PROGRAM ControlFBD
VAR
	qxLampStarted	AT %Q* : BOOL;
	qxSliderAout 	AT %Q* : BOOL; 
	qxSliderAin 	AT %Q* : BOOL; 
	qxSliderBout 	AT %Q* : BOOL; 
	qxSliderBin 	AT %Q* : BOOL; 
	qxDrillDown 	AT %Q* : BOOL;
	qxDrillUp		AT %Q* : BOOL;
	qxLampEmStopOk	AT %Q* : BOOL;
	qxLampSafetyOk  AT %Q* : BOOL;
	qxLampHomePos   AT %Q* : BOOL;
	
	
	mxManualRun : BOOL;
	mxEmergencyButtonPressed: BOOL;
	mxAuto : BOOL;
	mxAutoAIn : BOOL;
	mxAutoAOut : BOOL;
	mxAutoBIn : BOOL;
	mxAutoBOut : BOOL;
	mxAutoDrillDown: BOOL;
	mxAutoDrillUp: BOOL;
	
	mxSafetyOK : BOOL;
	mxManualOk : BOOL;
	mxCycleStopActivated : BOOL;
	mxBlink : BOOL;
	
	fbBlink : BLINK;

	
	
	ixButtonStart	AT %I* : BOOL;
	ixButtonStop	AT %I* : BOOL;
	ixSliderAout	AT %I* : BOOL;
	ixSliderAin		AT %I* : BOOL;
	ixSliderBout	AT %I* : BOOL;
	ixSliderBin		AT %I* : BOOL;
	ixDrillUp		AT %I* : BOOL;
	ixDrillDown		AT %I* : BOOL;

	ixAuto			AT %I* : BOOL;
	ixBtn1EmStopOk	AT %I* : BOOL;
	ixBtn2EmStopOk	AT %I* : BOOL;	
	ixSafety1StopOk	AT %I* : BOOL;
	ixSafety2StopOk	AT %I* : BOOL;	
	ixBtnReset		AT %I* : BOOL;
	ixBtnAout		AT %I* : BOOL;
	ixBtnAin		AT %I* : BOOL;
	ixBtnBout		AT %I* : BOOL;
	ixBtnBin		AT %I* : BOOL;
	ixBtnDrillOut	AT %I* : BOOL;
	ixBtnDrillIn	AT %I* : BOOL;

	mx: BOOL;
	mxStart: BOOL;
END_VAR

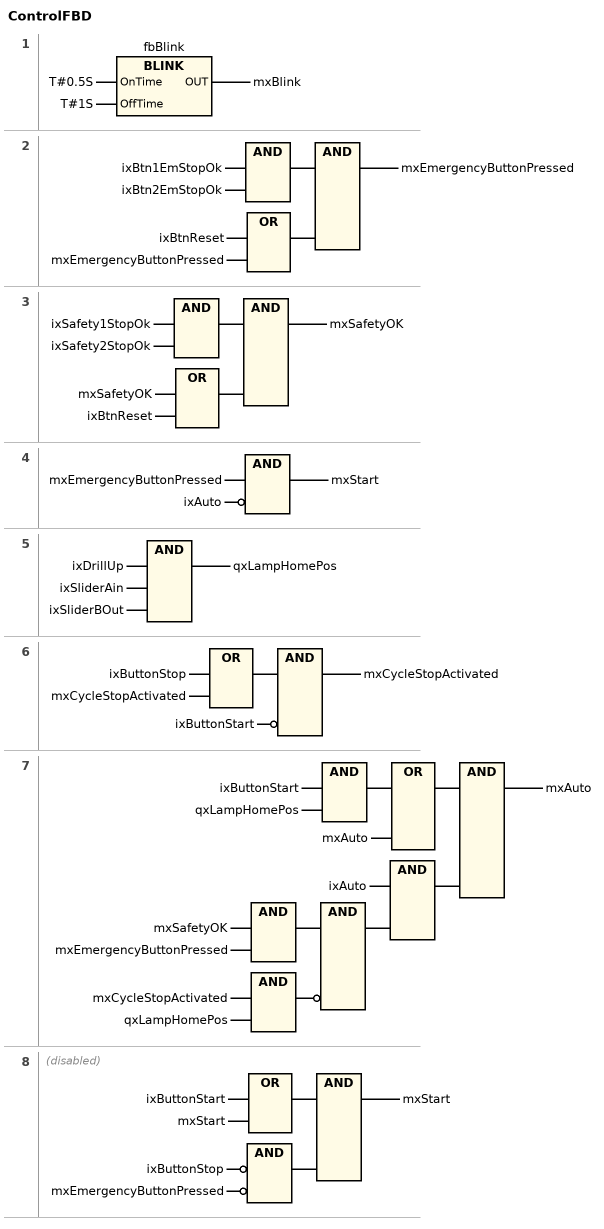
// NETWORK 1
fbBlink(OnTime := T#0.5S, OffTime := T#1S); // BLINK
mxBlink := fbBlink.OUT;

// NETWORK 2
mxEmergencyButtonPressed := (ixBtn1EmStopOk AND ixBtn2EmStopOk) AND (ixBtnReset OR mxEmergencyButtonPressed);

// NETWORK 3
mxSafetyOK := (ixSafety1StopOk AND ixSafety2StopOk) AND (mxSafetyOK OR ixBtnReset);

// NETWORK 4
mxStart := mxEmergencyButtonPressed AND NOT ixAuto;

// NETWORK 5
qxLampHomePos := ixDrillUp AND ixSliderAin AND ixSliderBOut;

// NETWORK 6
mxCycleStopActivated := (ixButtonStop OR mxCycleStopActivated) AND NOT ixButtonStart;

// NETWORK 7
mxAuto := (ixButtonStart AND qxLampHomePos OR mxAuto) AND (ixAuto AND ((mxSafetyOK AND mxEmergencyButtonPressed) AND NOT (mxCycleStopActivated AND qxLampHomePos)));

// NETWORK 8 (disabled)
// mxStart := (ixButtonStart OR mxStart) AND (NOT ixButtonStop AND NOT mxEmergencyButtonPressed);

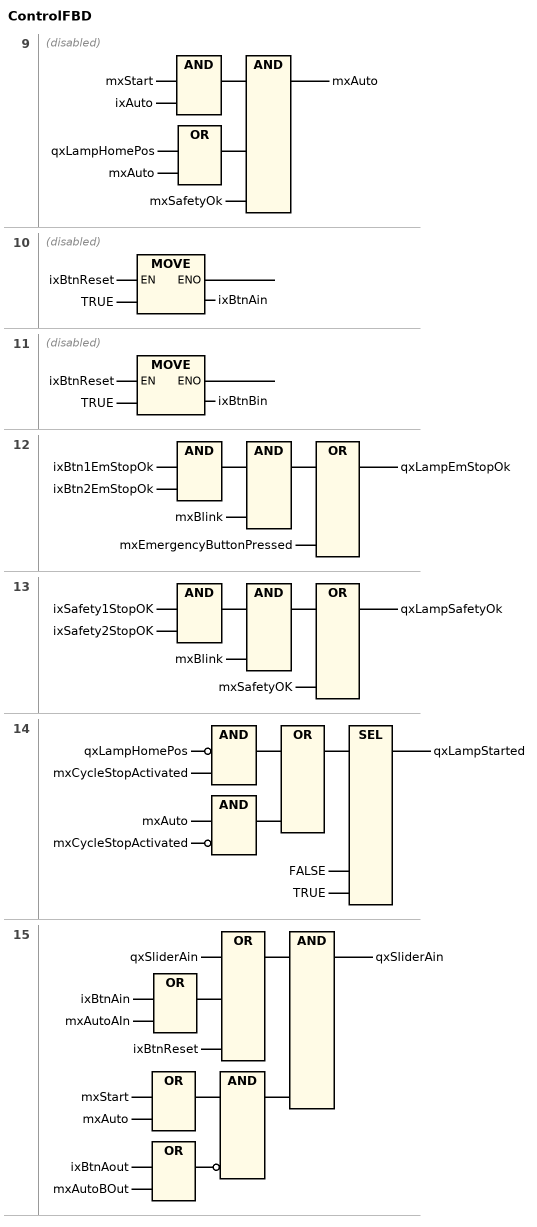
// NETWORK 9 (disabled)
// mxAuto := (mxStart AND ixAuto) AND (qxLampHomePos OR mxAuto) AND mxSafetyOk;

// NETWORK 10 (disabled)
// IF ixBtnReset THEN ixBtnAin := TRUE; END_IF

// NETWORK 11 (disabled)
// IF ixBtnReset THEN ixBtnBin := TRUE; END_IF

// NETWORK 12
qxLampEmStopOk := (ixBtn1EmStopOk AND ixBtn2EmStopOk) AND mxBlink OR mxEmergencyButtonPressed;

// NETWORK 13
qxLampSafetyOk := (ixSafety1StopOK AND ixSafety2StopOK) AND mxBlink OR mxSafetyOK;

// NETWORK 14
qxLampStarted := SEL(NOT qxLampHomePos AND mxCycleStopActivated OR mxAuto AND NOT mxCycleStopActivated, FALSE, TRUE);

// NETWORK 15
qxSliderAin := (qxSliderAin OR (ixBtnAin OR mxAutoAIn) OR ixBtnReset) AND ((mxStart OR mxAuto) AND NOT (ixBtnAout OR mxAutoBOut));

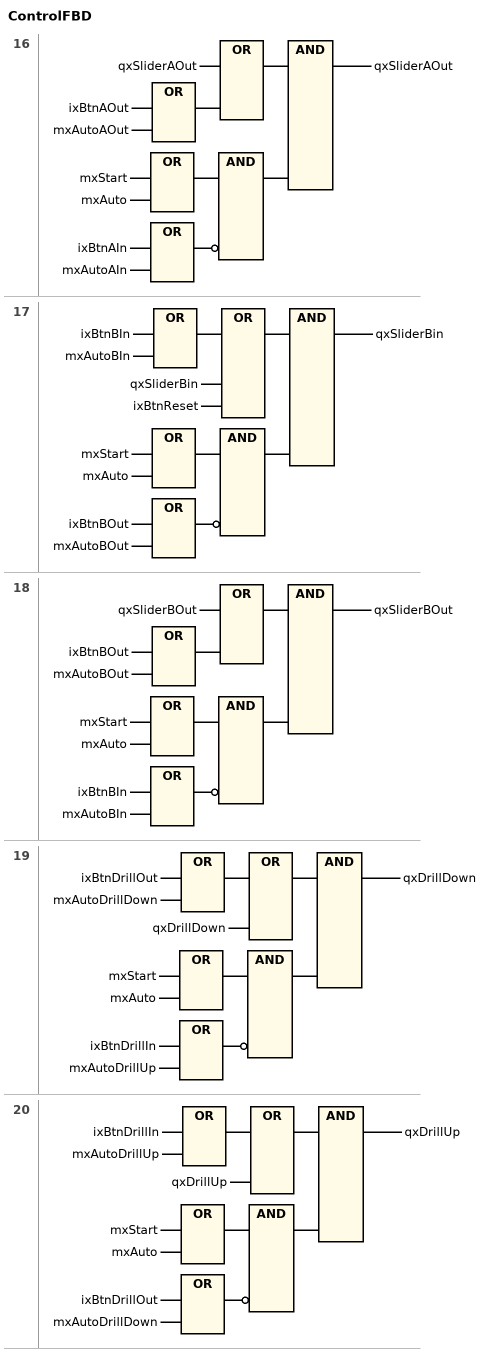
// NETWORK 16
qxSliderAOut := (qxSliderAOut OR (ixBtnAOut OR mxAutoAOut)) AND ((mxStart OR mxAuto) AND NOT (ixBtnAIn OR mxAutoAIn));

// NETWORK 17
qxSliderBin := ((ixBtnBIn OR mxAutoBIn) OR qxSliderBin OR ixBtnReset) AND ((mxStart OR mxAuto) AND NOT (ixBtnBOut OR mxAutoBOut));

// NETWORK 18
qxSliderBOut := (qxSliderBOut OR (ixBtnBOut OR mxAutoBOut)) AND ((mxStart OR mxAuto) AND NOT (ixBtnBIn OR mxAutoBIn));

// NETWORK 19
qxDrillDown := ((ixBtnDrillOut OR mxAutoDrillDown) OR qxDrillDown) AND ((mxStart OR mxAuto) AND NOT (ixBtnDrillIn OR mxAutoDrillUp));

// NETWORK 20
qxDrillUp := ((ixBtnDrillIn OR mxAutoDrillUp) OR qxDrillUp) AND ((mxStart OR mxAuto) AND NOT (ixBtnDrillOut OR mxAutoDrillDown));

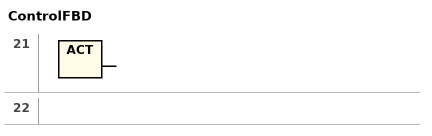
// NETWORK 21
ACT();

// NETWORK 22

ACTION ACT:
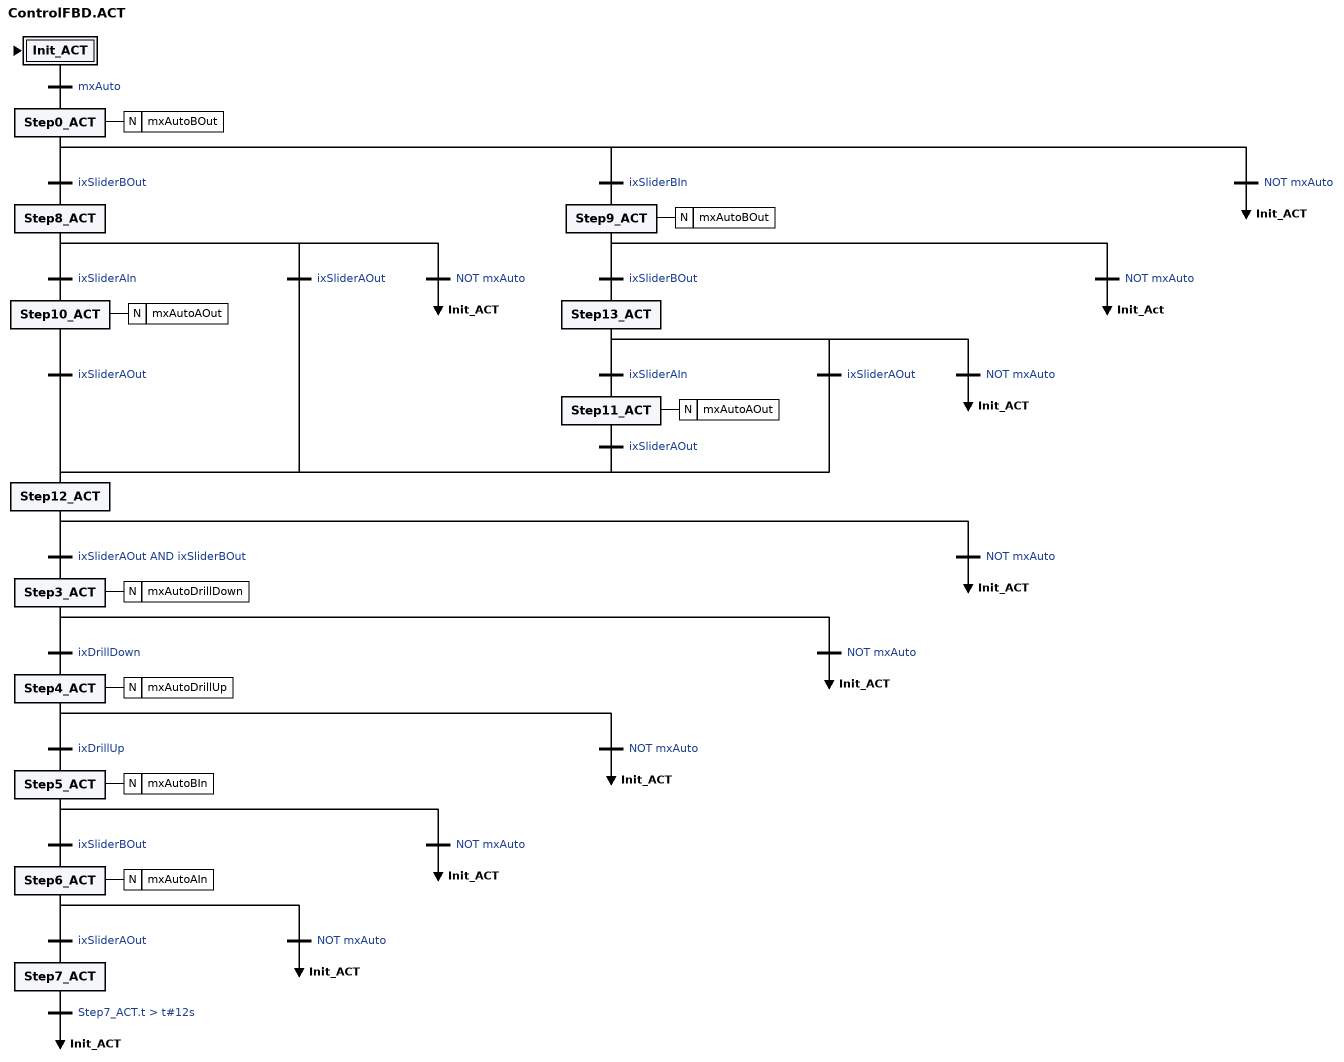
INITIAL_STEP Init_ACT:
END_STEP
TRANSITION FROM Init_ACT TO Step0_ACT
    := mxAuto;
END_TRANSITION
STEP Step0_ACT:
    mxAutoBOut(N);
END_STEP
TRANSITION FROM Step0_ACT TO Step8_ACT
    := ixSliderBOut;
END_TRANSITION
STEP Step8_ACT:
END_STEP
TRANSITION FROM Step8_ACT TO Step10_ACT
    := ixSliderAIn;
END_TRANSITION
STEP Step10_ACT:
    mxAutoAOut(N);
END_STEP
TRANSITION FROM Step10_ACT TO Step12_ACT
    := ixSliderAOut;
END_TRANSITION
TRANSITION FROM Step8_ACT TO Step12_ACT
    := ixSliderAOut;
END_TRANSITION
TRANSITION FROM Step8_ACT TO Init_ACT
    := NOT mxAuto;
END_TRANSITION
TRANSITION FROM Step0_ACT TO Step9_ACT
    := ixSliderBIn;
END_TRANSITION
STEP Step9_ACT:
    mxAutoBOut(N);
END_STEP
TRANSITION FROM Step9_ACT TO Step13_ACT
    := ixSliderBOut;
END_TRANSITION
TRANSITION FROM Step9_ACT TO Init_Act
    := NOT mxAuto;
END_TRANSITION
STEP Step13_ACT:
END_STEP
TRANSITION FROM Step13_ACT TO Step11_ACT
    := ixSliderAIn;
END_TRANSITION
STEP Step11_ACT:
    mxAutoAOut(N);
END_STEP
TRANSITION FROM Step11_ACT TO Step12_ACT
    := ixSliderAOut;
END_TRANSITION
TRANSITION FROM Step13_ACT TO Step12_ACT
    := ixSliderAOut;
END_TRANSITION
TRANSITION FROM Step13_ACT TO Init_ACT
    := NOT mxAuto;
END_TRANSITION
TRANSITION FROM Step0_ACT TO Init_ACT
    := NOT mxAuto;
END_TRANSITION
STEP Step12_ACT:
END_STEP
TRANSITION FROM Step12_ACT TO Step3_ACT
    := ixSliderAOut AND ixSliderBOut;
END_TRANSITION
TRANSITION FROM Step12_ACT TO Init_ACT
    := NOT mxAuto;
END_TRANSITION
STEP Step3_ACT:
    mxAutoDrillDown(N);
END_STEP
TRANSITION FROM Step3_ACT TO Step4_ACT
    := ixDrillDown;
END_TRANSITION
TRANSITION FROM Step3_ACT TO Init_ACT
    := NOT mxAuto;
END_TRANSITION
STEP Step4_ACT:
    mxAutoDrillUp(N);
END_STEP
TRANSITION FROM Step4_ACT TO Step5_ACT
    := ixDrillUp;
END_TRANSITION
TRANSITION FROM Step4_ACT TO Init_ACT
    := NOT mxAuto;
END_TRANSITION
STEP Step5_ACT:
    mxAutoBIn(N);
END_STEP
TRANSITION FROM Step5_ACT TO Step6_ACT
    := ixSliderBOut;
END_TRANSITION
TRANSITION FROM Step5_ACT TO Init_ACT
    := NOT mxAuto;
END_TRANSITION
STEP Step6_ACT:
    mxAutoAIn(N);
END_STEP
TRANSITION FROM Step6_ACT TO Step7_ACT
    := ixSliderAOut;
END_TRANSITION
TRANSITION FROM Step6_ACT TO Init_ACT
    := NOT mxAuto;
END_TRANSITION
STEP Step7_ACT:
END_STEP
TRANSITION FROM Step7_ACT TO Init_ACT
    := Step7_ACT.t > t#12s;
END_TRANSITION
// branch label Branch1_ACT
// branch label Branch3_ACT
// branch label Branch2_ACT
// branch label Branch0_ACT
// branch label Branch4_ACT
// branch label Branch5_ACT
// branch label Branch6_ACT
// branch label Branch7_ACT
// branch label Branch8_ACT
END_ACTION

ACTION Step14_ACT_exit:

END_ACTION

END_PROGRAM

(* stored: Version 1.1.0.1
   POU ControlFBD: Id {441bf843-2f16-42db-a10b-d561aec11b1f}, SpecialFunc None
   Action ACT: Id {f91e217c-2f17-48ef-ae7e-14449dcdbd88}
   Action Step14_ACT_exit: Id {c5ba0539-4636-4576-887c-1fcac97cd435} *)
